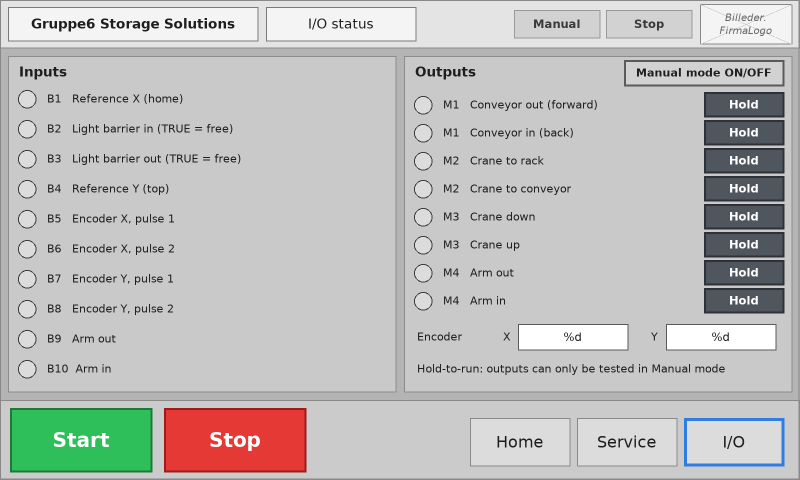
VISUALIZATION IO  // 800x480
    Rectangle (0,0 800x480)
    Rectangle (0,0 800x48)
    Rectangle (8,7 250x34), "Gruppe6 Storage Solutions"
    Rectangle (266,7 150x34), "I/O status"
    Rectangle (514,10 86x28), "Manual", colour toggle: MAIN.isManualMode
    Rectangle (606,10 86x28), "Stop", colour toggle: MAIN.isStop
    Image (700,4 92x40), image: Billeder.FirmaLogo
    Rectangle (0,400 800x80)
    RoundedRectangle (10,408 142x64), "Start"
        OnMouseUp: execute { MAIN.isStop := FALSE; }
    RoundedRectangle (164,408 142x64), "Stop"
        OnMouseUp: execute { MAIN.isStop := TRUE; }
    Rectangle (470,418 100x48), "Home"
        OnMouseUp: execute {
            MAIN.logoutRequest := TRUE;   // leaving the service page logs out
        }
        OnMouseUp: change screen: Start
    Rectangle (577,418 100x48), "Service"
        OnMouseUp: change screen: Service
    Rectangle (684,418 100x48), "I/O"
    Rectangle (8,56 388x336)
    Rectangle (16,60 372x24), "Inputs"
    Ellipse (18,90 18x18), colour toggle: MAIN.B1
    Rectangle (44,86 330x26), "B1 Reference X (home)"
    Ellipse (18,120 18x18), colour toggle: MAIN.B2
    Rectangle (44,116 330x26), "B2 Light barrier in (TRUE = free)"
    Ellipse (18,150 18x18), colour toggle: MAIN.B3
    Rectangle (44,146 330x26), "B3 Light barrier out (TRUE = free)"
    Ellipse (18,180 18x18), colour toggle: MAIN.B4
    Rectangle (44,176 330x26), "B4 Reference Y (top)"
    Ellipse (18,210 18x18), colour toggle: MAIN.B5
    Rectangle (44,206 330x26), "B5 Encoder X, pulse 1"
    Ellipse (18,240 18x18), colour toggle: MAIN.B6
    Rectangle (44,236 330x26), "B6 Encoder X, pulse 2"
    Ellipse (18,270 18x18), colour toggle: MAIN.B7
    Rectangle (44,266 330x26), "B7 Encoder Y, pulse 1"
    Ellipse (18,300 18x18), colour toggle: MAIN.B8
    Rectangle (44,296 330x26), "B8 Encoder Y, pulse 2"
    Ellipse (18,330 18x18), colour toggle: MAIN.B9
    Rectangle (44,326 330x26), "B9 Arm out"
    Ellipse (18,360 18x18), colour toggle: MAIN.B10
    Rectangle (44,356 330x26), "B10 Arm in"
    Rectangle (404,56 388x336)
    Rectangle (412,60 372x24), "Outputs"
    RoundedRectangle (624,60 160x26), "Manual mode ON/OFF", colour toggle: MAIN.isManualMode
        toggle MAIN.isManualMode
    Ellipse (414,96 18x18), colour toggle: MAIN.M1_Forward
    Rectangle (440,92 250x26), "M1 Conveyor out (forward)"
    RoundedRectangle (704,92 80x25), "Hold", input disabled if: MAIN.ioTestLocked
        tap MAIN.testM1Forward
    Ellipse (414,124 18x18), colour toggle: MAIN.M1_Back
    Rectangle (440,120 250x26), "M1 Conveyor in (back)"
    RoundedRectangle (704,120 80x25), "Hold", input disabled if: MAIN.ioTestLocked
        tap MAIN.testM1Back
    Ellipse (414,152 18x18), colour toggle: MAIN.M2_Forward
    Rectangle (440,148 250x26), "M2 Crane to rack"
    RoundedRectangle (704,148 80x25), "Hold", input disabled if: MAIN.ioTestLocked
        tap MAIN.testM2Forward
    Ellipse (414,180 18x18), colour toggle: MAIN.M2_Back
    Rectangle (440,176 250x26), "M2 Crane to conveyor"
    RoundedRectangle (704,176 80x25), "Hold", input disabled if: MAIN.ioTestLocked
        tap MAIN.testM2Back
    Ellipse (414,208 18x18), colour toggle: MAIN.M3_Down
    Rectangle (440,204 250x26), "M3 Crane down"
    RoundedRectangle (704,204 80x25), "Hold", input disabled if: MAIN.ioTestLocked
        tap MAIN.testM3Down
    Ellipse (414,236 18x18), colour toggle: MAIN.M3_Up
    Rectangle (440,232 250x26), "M3 Crane up"
    RoundedRectangle (704,232 80x25), "Hold", input disabled if: MAIN.ioTestLocked
        tap MAIN.testM3Up
    Ellipse (414,264 18x18), colour toggle: MAIN.M4_Forward
    Rectangle (440,260 250x26), "M4 Arm out"
    RoundedRectangle (704,260 80x25), "Hold", input disabled if: MAIN.ioTestLocked
        tap MAIN.testM4Forward
    Ellipse (414,292 18x18), colour toggle: MAIN.M4_Back
    Rectangle (440,288 250x26), "M4 Arm in"
    RoundedRectangle (704,288 80x25), "Hold", input disabled if: MAIN.ioTestLocked
        tap MAIN.testM4Back
    Rectangle (414,324 80x26), "Encoder"
    Rectangle (500,324 20x26), "X"
    Rectangle (518,324 110x26), "%d", text variable: MAIN.currentPosX
    Rectangle (648,324 20x26), "Y"
    Rectangle (666,324 110x26), "%d", text variable: MAIN.currentPosY
    Rectangle (414,356 370x26), "Hold-to-run: outputs can only be tested in Manual mode"
END_VISUALIZATION

(* stored: Version 1.1.0.1, ProductVersion 3.1.4024.12
   Visu IO: Id {8da2a5a5-256d-4ba0-861e-2393506b703d} *)
